// TIA Portal V21 export
// export: Created 2026-11-10T19:21:31.5036988Z, ExportSetting WithDefaults, DisplayName Totally Integrated Automation Portal, DisplayVersion V21 Update 3, DisplayName STEP 7 Professional, DisplayVersion V21 Update 3, DisplayName STEP 7 Safety, DisplayVersion V21, DisplayName Tech WebApplication, DisplayVersion V21, DisplayName WinCC Basic/Comfort/Advanced, DisplayVersion V21 Update 3, DisplayName WinCC Unified, DisplayVersion V21 Update 3
FUNCTION_BLOCK "FB_Lad_mb001"   // FB5, LAD
{ S7_Optimized_Access := 'TRUE' }
VERSION : 0.1
// stored: AutoNumber true, IsIECCheckEnabled false, IsRetainMemResEnabled false, MemoryReserve 100, SetENOAutomatically false, UDAEnableTagReadback false
   VAR_INPUT
      v_req : Bool;
      v_port : PORT;
      v_baud : UDInt;
      v_parity : UInt;
      v_flow_ctrl : UInt;
      v_rts_on_dly : UInt;
      v_rts_off_dly : UInt;
      v_resp_to : UInt;
   END_VAR
   VAR_OUTPUT
      v_done : Bool;
      v_error : Bool;
      v_status : Word;
   END_VAR
   VAR_IN_OUT
      v_mb_db : P2P_MB_BASE;
   END_VAR
   VAR
      inst { S7_SetPoint := 'True'} : Modbus_Comm_Load;
   END_VAR
BEGIN

REGION Network 1: MB_COMM_LOAD - Configure port on the PtP module for Modbus RTU
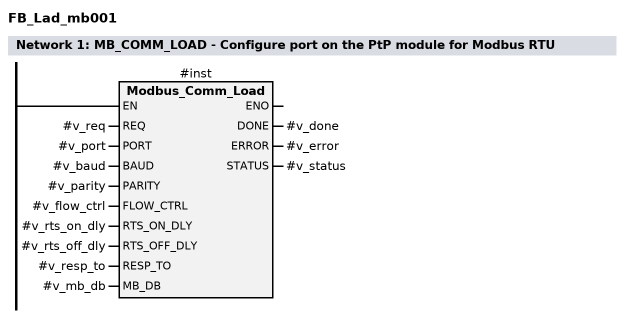
   RUNG wire#powerrail
      #inst.Modbus_Comm_Load(REQ := #v_req, PORT := #v_port, BAUD := #v_baud, PARITY := #v_parity, FLOW_CTRL := #v_flow_ctrl, RTS_ON_DLY := #v_rts_on_dly, RTS_OFF_DLY := #v_rts_off_dly, RESP_TO := #v_resp_to, MB_DB := #v_mb_db, DONE => #v_done, ERROR => #v_error, STATUS => #v_status)
   END_RUNG
   // the same network as SCL:
   #inst(REQ := #v_req,   // Modbus_Comm_Load
         PORT := #v_port,
         BAUD := #v_baud,
         PARITY := #v_parity,
         FLOW_CTRL := #v_flow_ctrl,
         RTS_ON_DLY := #v_rts_on_dly,
         RTS_OFF_DLY := #v_rts_off_dly,
         RESP_TO := #v_resp_to,
         MB_DB := #v_mb_db,
         DONE => #v_done,
         ERROR => #v_error,
         STATUS => #v_status);
END_REGION
END_FUNCTION_BLOCK
